// TIA Portal V21 export
// export: Created 2026-11-08T19:47:34.5615124Z, ExportSetting WithDefaults, DisplayName Totally Integrated Automation Portal, DisplayVersion V21 Update 3, DisplayName STEP 7 Professional, DisplayVersion V21 Update 3, DisplayName STEP 7 Safety, DisplayVersion V21, DisplayName Tech WebApplication, DisplayVersion V21, DisplayName WinCC Basic/Comfort/Advanced, DisplayVersion V21 Update 3, DisplayName WinCC Unified, DisplayVersion V21 Update 3
FUNCTION "FC_Scl" : Void   // FC1, SCL
{ S7_Optimized_Access := 'TRUE' }
VERSION : 0.1
// stored: AutoNumber true, IsIECCheckEnabled false, SetENOAutomatically false, UDAEnableTagReadback false
   VAR_INPUT
      "a" : Int;   // First input
      "b" : Int;   // Second input
   END_VAR
   VAR_OUTPUT
      result : Int;   // Limited sum
      total : Int;   // Sum 1..4
   END_VAR
   VAR_IN_OUT
      gain : Real;   // Gain value
   END_VAR
   VAR_TEMP
      tmp : Int;
      i : Int;
   END_VAR
BEGIN
   // Sum of both inputs
   #tmp := #a + #b;

   // Limit the result to 0..100
   #result := 0;
   IF #tmp > 100 THEN
       #result := 100;
   ELSIF #tmp < 0 THEN
       #result := 0;
   ELSE
       #result := #tmp;
   END_IF;

   // Accumulate 1..4
   #total := 0;
   FOR #i := 1 TO 4 DO
       #total := #total + #i;
   END_FOR;

   // Call the function block with its instance data block
   "FB_Iface_DB"(iBool := TRUE,
                 iInt := #result,
                 iReal := 1.5,
                 ioReal := #gain);
END_FUNCTION
